Staubli VAL3: action_do.pgx

public program action_do(num x_nIndex)
  local num l_nType
  local string l_sType
  local bool l_bActive
  local string l_sBoolValue
  local num l_nBoolValue
  local num l_nIOindex
  local num l_nPulseValue
  local num l_i
begin
  for l_i = 0 to size(actionData:aActItem[x_nIndex].aActItem)-1
    l_sType=actionData:aActItem[x_nIndex].aActItem[l_i].sIOtype
    l_bActive=(actionData:aActItem[x_nIndex].aActItem[l_i].bActive==true)
    l_sBoolValue=actionData:aActItem[x_nIndex].aActItem[l_i].sValue
    l_nIOindex=actionData:aActItem[x_nIndex].aActItem[l_i].nIOindex
    l_nPulseValue=actionData:aActItem[x_nIndex].aActItem[l_i].nPulseValue
    switch l_sBoolValue
      case "ON"
        l_nBoolValue=1
      break
      case "OFF"
        l_nBoolValue=0
      break
    endSwitch
    if l_bActive
      switch l_sType
        case "IN"
          call addActCmd(1,3,l_nIOindex,l_nBoolValue)
        break
        case "OUT"
          call addActCmd(1,1,l_nIOindex,l_nBoolValue)
        break
        case "PULSE"
          call addActCmd(1,2,l_nIOindex,l_nPulseValue)
        break

      endSwitch
    endIf
  endFor
  popUpMsg("执行动作："+toString("",x_nIndex))
end
